(* IEC 61131-3 sources: rusty/tests/lit/single/complex_return_types, 5 files *)

(* ---- array_of_array_returns.st ---- *)
// RUN: %COMPILE %s && %RUN | %CHECK %s
// XFAIL: *
// Fails because of #1389
FUNCTION foo : ARRAY[0..1] OF ARRAY[0..1] OF INT
    VAR
        result : ARRAY[0..1] OF ARRAY[0..1] OF INT;
    END_VAR
    result[0][0] := 5;
    result[0][1] := 10;
    result[1][0] := 15;
    result[1][1] := 20;
    foo := result;
END_FUNCTION

FUNCTION bar : ARRAY[0..1] OF ARRAY[0..1] OF INT
    VAR
        data : ARRAY[0..1] OF ARRAY[0..1] OF INT;
    END_VAR
    data := foo();
    bar := data;
END_FUNCTION

FUNCTION baz : ARRAY[0..2] OF STRING[20]
    VAR
        texts : ARRAY[0..2] OF STRING[20];
    END_VAR
    texts[0] := 'One';
    texts[1] := 'Two';
    texts[2] := 'Three';
    baz := texts;
END_FUNCTION

FUNCTION main
    VAR
        numbers : ARRAY[0..1] OF ARRAY[0..1] OF INT;
        strings : ARRAY[0..2] OF STRING[20];
    END_VAR
    numbers := bar();
    strings := baz();

    // CHECK: 5 10 15 20
    printf('%d %d %d %d$N', numbers[0][0], numbers[0][1], numbers[1][0], numbers[1][1]);

    // CHECK: One Two Three
    printf('%s %s %s$N', REF(strings[0]), REF(strings[1]), REF(strings[2]));
END_FUNCTION

(* ---- array_of_string_return.st ---- *)
// RUN: %COMPILE %s && %RUN | %CHECK %s
// XFAIL: *
// Fails because of #1389
FUNCTION func_with_aggregagte_return: ARRAY[0..1] OF STRING
VAR_INPUT
    in: STRING;
    in2: STRING;
END_VAR
    func_with_aggregagte_return[0] := in;
    func_with_aggregagte_return[1] := in2;
END_FUNCTION

FUNCTION main : DINT
VAR
    ret : ARRAY[0..1] OF STRING;
END_VAR
    ret := func_with_aggregagte_return('Hello', 'World!');
    printf('%s$N', ADR(ret[0])); //CHECK Hello
    printf('%s$N', ADR(ret[1])); //CHECK World!
END_FUNCTION

(* ---- function_with_explicit_calls.st ---- *)
// RUN: %COMPILE %s && %RUN | %CHECK %s
FUNCTION foo : STRING
        VAR_INPUT
            x : DINT;
        END_VAR
        foo := 'hello';
END_FUNCTION
FUNCTION main : DINT
VAR
    res : STRING;
END_VAR
    res := foo(x := 1);
    printf('%s$N', ADR(res)); // CHECK: hello
END_FUNCTION

(* ---- nested_string_return_call_in_if_condition.st ---- *)
// RUN: %COMPILE %s && %RUN | %CHECK %s
FUNCTION CLEAN : STRING
VAR_INPUT
    IN : STRING;
	CX : STRING;
END_VAR
VAR
	pos: INT := 1;
    stop: INT;
END_VAR
    CLEAN := IN;
    stop := LEN(IN);
    WHILE pos <= stop DO
        IF FIND(CX, MID(CLEAN, 1, pos)) > 0 THEN
            pos := pos + 1;
        ELSE
            CLEAN := DELETE(CLEAN, 1, pos);
            stop := stop - 1;
        END_IF;
    END_WHILE;
END_FUNCTION

FUNCTION main : DINT
VAR
    needle: STRING := 'aeiou ,?';
    haystack: STRING := 'hello world, how are you?';
    result: STRING;
END_VAR
    result := CLEAN(haystack, needle);
    printf('%s$N', REF(result)); // CHECK: eo o, o ae ou?
END_FUNCTION

(* ---- string_return_function_called_in_while_loop.st ---- *)
// RUN: %COMPILE %s && %RUN | %CHECK %s
FUNCTION TRIM : STRING
VAR_INPUT
	str : STRING;
END_VAR

TRIM := str;
WHILE LEFT(TRIM, 1) = ' ' DO
	TRIM := DELETE(TRIM, 1, 1);
END_WHILE;

IF RIGHT(TRIM, 1) = ' ' THEN
REPEAT
	TRIM := DELETE(TRIM, 1, LEN(TRIM));
UNTIL RIGHT(TRIM, 1) <> ' '
END_REPEAT;
END_IF;

END_FUNCTION

FUNCTION main
VAR
    str : STRING := '  hello world  ';
END_VAR
    printf('%s$N', REF(TRIM(str))); // CHECK: hello world
END_FUNCTION
